// TIA Portal V21 export
// export: Created 2026-10-12T12:46:18.9630019Z, ExportSetting WithDefaults, DisplayName Totally Integrated Automation Portal, DisplayVersion V21, DisplayName STEP 7 Professional, DisplayVersion V21, DisplayName STEP 7 Safety, DisplayVersion V21, DisplayName Tech WebApplication, DisplayVersion V21, DisplayName WinCC Basic/Comfort/Advanced, DisplayVersion V21, DisplayName WinCC Unified, DisplayVersion V21
TagTable "ALARMS"
  ALARM WORD : Int  (%DB2.DBW0, HMI_Connection_1, 1 s)
